TYPE ST_MachinePermissives :
STRUCT
    bSafetyIndexPermissive   : BOOL;
    bOperatorIndexPermissive : BOOL;
    bStationsIndexPermissive : BOOL;
    bIndexMoveAllowed        : BOOL;
    bAirSupplyReady          : BOOL;
    bDoorInitialisationReady : BOOL;
    bIndexInitialisationReady: BOOL;
    bStationsHome            : BOOL;
    bInitialisationAllowed   : BOOL;
    bAutoCycleAllowed        : BOOL;
END_STRUCT
END_TYPE

(* stored: Version 1.1.0.1, ProductVersion 3.1.4026.18
   DUT ST_MachinePermissives: Id {c1eb91aa-e552-4751-9960-a96c109c7f62} *)
